Staubli VAL3: getMoveType.pgx

public program getMoveType(string x_sKey, num x_nIndex, num& x_nMoveType)
begin
  x_nMoveType=trajTemp:tTrajItem[x_sKey].pPointItem[x_nIndex].pParaItem.nMoveType
end
